(* IEC 61131-3 sources: SRCI_CLIENT_PLC/RobotLibrary/Library/Structures/Data/WorkArea, 4 files *)

(* ---- RobotWorkArea.st ---- *)
{attribute 'pack_mode' := '1'}
// -------------------------------------------------------------------------
//  SRCI Robot Library
// -------------------------------------------------------------------------
//
//  Object:      RobotWorkArea
//  Author:      Thorsten Brach
//  Date:        2025-04-22
//
//  Description:
//
//
//  Copyright:
//    (C) 2025 Thorsten Brach. All rights reserved
//             Licensed under the MIT License.
//
//  Disclaimer:
//    This project is provided without any guarantee and can be used for
//    private and commercial purposes. Any use is at the user’s
//    own risk and responsibility.
//
// -------------------------------------------------------------------------
TYPE RobotWorkArea :
STRUCT
  /// Workarea is available
  Available : BOOL;
  /// Workarea data
  Data      : RobotWorkAreaData;
END_STRUCT
END_TYPE

(* ---- RobotWorkAreaData.st ---- *)
{attribute 'pack_mode' := '1'}
// -------------------------------------------------------------------------
//  SRCI Robot Library
// -------------------------------------------------------------------------
//
//  Object:      RobotWorkAreaData
//  Author:      Thorsten Brach
//  Date:        2024-06-01
//
//  Description:
//
//
//  Copyright:
//    (C) 2024 Thorsten Brach. All rights reserved
//             Licensed under the MIT License.
//
//  Disclaimer:
//    This project is provided without any guarantee and can be used for
//    private and commercial purposes. Any use is at the user’s
//    own risk and responsibility.
//
// -------------------------------------------------------------------------
TYPE RobotWorkAreaData :
STRUCT
  /// Timestamp
  Timestamp          : IEC_TIMESTAMP;
  /// Defines type of work area
  AreaType           : AreaType := AreaTypeEnum.BOX; // ST-FIX F156: spec 5.5.8 table 5-34: 1 Box (default); alias AreaTypeEnum because the member has the name of the type
  /// Defines violation condition
  /// • FALSE (default) : Robot must not leave defined area
  /// • TRUE            : Robot must not enter defined area
  AreaMode           : BOOL := FALSE;
  /// Defines RC’s and robot’s behavior when robot violates work area
  ReactionMode       : WorkAreaReactionMode;
  /// Specifies whether an active work area can be edited by function WriteWorkArea
  ///  TRUE            : Modification of active work area possible
  ///  FALSE (default) : Modification of active work areas not possible
  ActiveModification : BOOL;
  /// Relates to AreaType Box, Cylinder and Sphere.
  DefinitionMode     : DefinitionMode;
  /// Relates to AreaType Box, Cylinder and Sphere.
  /// Index of reference frame
  /// • 0: WCS (default)
  /// • 1..254: User frames
  FrameNo            : USINT;
  /// Relates to AreaType Box, Cylinder and Sphere.
  /// X-value of reference point in specified frame - Default: 0
  ZeroPointX         : REAL := 0;
  /// Relates to AreaType Box, Cylinder and Sphere.
  /// Y-value of reference point in specified frame - Default: 0
  ZeroPointY         : REAL := 0;
  /// Relates to AreaType Box, Cylinder and Sphere.
  /// Z-value of reference point in specified frame - Default: 0
  ZeroPointZ         : REAL := 0;
  /// Limit for cartesian X
  X                  : RobotWorkAreaDataLimitCartesian;
  /// Limit for cartesian Y
  Y                  : RobotWorkAreaDataLimitCartesian;
  /// Limit for cartesian Z
  Z                  : RobotWorkAreaDataLimitCartesian;
  /// Relates to AreaType Sphere.
  /// Radius of cylinder or sphere - Default 0
  Radius             : REAL := 0;
  /// Limits for Joint J1
  J1Limit            : RobotWorkAreaDataLimitJoint;
  /// Limits for Joint J2
  J2Limit            : RobotWorkAreaDataLimitJoint;
  /// Limits for Joint J3
  J3Limit            : RobotWorkAreaDataLimitJoint;
  /// Limits for Joint J4
  J4Limit            : RobotWorkAreaDataLimitJoint;
  /// Limits for Joint J5
  J5Limit            : RobotWorkAreaDataLimitJoint;
  /// Limits for Joint J6
  J6Limit            : RobotWorkAreaDataLimitJoint;
  /// Limits for Joint E1
  E1Limit            : RobotWorkAreaDataLimitJoint;
  /// Limits for Joint E2
  E2Limit            : RobotWorkAreaDataLimitJoint;
  /// Limits for Joint E3
  E3Limit            : RobotWorkAreaDataLimitJoint;
  /// Limits for Joint E4
  E4Limit            : RobotWorkAreaDataLimitJoint;
  /// Limits for Joint E5
  E5Limit            : RobotWorkAreaDataLimitJoint;
  /// Limits for Joint E6
  E6Limit            : RobotWorkAreaDataLimitJoint;
END_STRUCT
END_TYPE

(* ---- RobotWorkAreaDataLimitCartesian.st ---- *)
{attribute 'pack_mode' := '1'}
// -------------------------------------------------------------------------
//  SRCI Robot Library
// -------------------------------------------------------------------------
//
//  Object:      RobotWorkAreaDataLimitCartesian
//  Author:      Thorsten Brach
//  Date:        2024-06-01
//
//  Description:
//
//
//  Copyright:
//    (C) 2024 Thorsten Brach. All rights reserved
//             Licensed under the MIT License.
//
//  Disclaimer:
//    This project is provided without any guarantee and can be used for
//    private and commercial purposes. Any use is at the user’s
//    own risk and responsibility.
//
// -------------------------------------------------------------------------
TYPE RobotWorkAreaDataLimitCartesian :
STRUCT
  /// Relates to AreaType Box, Cylinder and Sphere.
  /// Distance in negative Direction - Default 0
  LowerLimit : REAL := 0;
  /// Relates to AreaType Box, Cylinder and Sphere.
  /// Distance in positive Direction - Default 0
  UpperLimit : REAL := 0;
END_STRUCT
END_TYPE

(* ---- RobotWorkAreaDataLimitJoint.st ---- *)
{attribute 'pack_mode' := '1'}
// -------------------------------------------------------------------------
//  SRCI Robot Library
// -------------------------------------------------------------------------
//
//  Object:      RobotWorkAreaDataLimitJoint
//  Author:      Thorsten Brach
//  Date:        2024-06-01
//
//  Description:
//
//
//  Copyright:
//    (C) 2024 Thorsten Brach. All rights reserved
//             Licensed under the MIT License.
//
//  Disclaimer:
//    This project is provided without any guarantee and can be used for
//    private and commercial purposes. Any use is at the user’s
//    own risk and responsibility.
//
// -------------------------------------------------------------------------
TYPE RobotWorkAreaDataLimitJoint :
STRUCT
  /// Relates to AreaType Axes.
  /// Negative work area limit for Joint
  /// • 0 (default) : No work area restriction of joint if lower and upper limit are set to 0
  /// • 16#FFFF_FFFF: No lower work area restrictions for Joint
  LowerLimit : REAL := 0;
  /// Relates to AreaType Axes.
  /// positive work area limit for Joint
  /// • 0 (default) : No work area restriction of joint if lower and upper limit of are set to 0
  /// • 16#FFFF_FFFF: No lower work area restrictions for Joint
  UpperLimit : REAL := 0;
END_STRUCT
END_TYPE
